FUNCTION_BLOCK SortingCycle_HMI (* Service Interface Function Block Type *)
  (* Standard: 61499-2 *)
  (* Version 0.0, 10/19/2026, sorting2n, Schneider Electric, template *)
  PACKAGE Main;
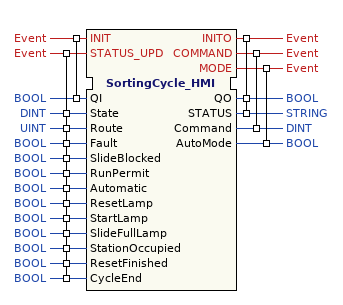
  EVENT_INPUT
    INIT WITH QI;
    STATUS_UPD WITH State, Route, Fault, SlideBlocked, RunPermit, Automatic, ResetLamp, StartLamp, SlideFullLamp, StationOccupied, ResetFinished, CycleEnd;
  END_EVENT
  EVENT_OUTPUT
    INITO WITH QO, STATUS;
    COMMAND WITH Command;
    MODE WITH AutoMode;
  END_EVENT
  VAR_INPUT
    QI : BOOL;
    State : DINT;
    Route : UINT;
    Fault : BOOL;
    SlideBlocked : BOOL;
    RunPermit : BOOL;
    Automatic : BOOL;
    ResetLamp : BOOL := FALSE;
    StartLamp : BOOL := FALSE;
    SlideFullLamp : BOOL := FALSE;
    StationOccupied : BOOL := FALSE;
    ResetFinished : BOOL := FALSE;
    CycleEnd : BOOL := FALSE;
  END_VAR
  VAR_OUTPUT
    QO : BOOL;
    STATUS : STRING;
    Command : DINT;
    AutoMode : BOOL;
  END_VAR
  SERVICE /
    SEQUENCE 
    END_SEQUENCE
  END_SERVICE
END_FUNCTION_BLOCK
